TYPE "DigValFF"
VERSION : 0.0
   STRUCT
      Value : Bool;   // Value
      InternalUseBit1 { ExternalAccessible := 'False'; ExternalVisible := 'False'; ExternalWritable := 'False'; CFC_Configurable := 'false'; CFC_Interconnectable := 'false'} : Bool;   // ByPass
      InternalUseBit2 { ExternalAccessible := 'False'; ExternalVisible := 'False'; ExternalWritable := 'False'; CFC_Configurable := 'false'; CFC_Interconnectable := 'false'} : Bool;   // Reserved
      InternalUseBit3 { ExternalAccessible := 'False'; ExternalVisible := 'False'; ExternalWritable := 'False'; CFC_Configurable := 'false'; CFC_Interconnectable := 'false'} : Bool;   // Reserved
      InternalUseBit4 { ExternalAccessible := 'False'; ExternalVisible := 'False'; ExternalWritable := 'False'; CFC_Configurable := 'false'; CFC_Interconnectable := 'false'} : Bool;   // Reserved
      InternalUseBit5 { ExternalAccessible := 'False'; ExternalVisible := 'False'; ExternalWritable := 'False'; CFC_Configurable := 'false'; CFC_Interconnectable := 'false'} : Bool;   // Reserved
      InternalUseBit6 { ExternalAccessible := 'False'; ExternalVisible := 'False'; ExternalWritable := 'False'; CFC_Configurable := 'false'; CFC_Interconnectable := 'false'} : Bool;   // Reserved
      InternalUseBit7 { ExternalAccessible := 'False'; ExternalVisible := 'False'; ExternalWritable := 'False'; CFC_Configurable := 'false'; CFC_Interconnectable := 'false'} : Bool;   // Reserved
      ST : Byte := BYTE#16#FF;   // Signal Status
   END_STRUCT;

END_TYPE

